(*
SPDX-FileCopyrightText: © 2026 Oleksandr Tiutyk <trofimich@gmail.com>
SPDX-License-Identifier: MIT
License: https://opensource.org/license/mit
*)

(*!
<summary>Orders WSTRING(255) values described by generic descriptors.</summary>
<description>
Non-null addresses must reference live WSTRING(255) storage. TypeClass and Size are not validated and no
numeric conversion is performed. Two null addresses compare equal; one null address sorts before a non-null
address. Uses native string comparison through the declared 255-character pointer type; descriptor Size does
not bound the read. Descriptors are passed by value; payload remains borrowed and is not modified, cloned,
released or retained. IsMemoryOwner does not affect comparison.
</description>
*)

FUNCTION_BLOCK WStringComparer EXTENDS TOF_Core.Object IMPLEMENTS TOF_Core.IComparer
VAR_STAT
	//! <summary>Class name shared by all instances of this function block.</summary>
	{attribute 'hide'} 
	_ClassName : STRING := __POUNAME();
END_VAR

{attribute 'monitoring' := 'call'}
PROPERTY ClassName : REFERENCE TO STRING
GET
ClassName REF= _ClassName;
END_GET
END_PROPERTY

(*!
<summary>Compares the first operand with the second using this ordering strategy.</summary>
<description>
Non-null addresses must reference live WSTRING(255) storage. TypeClass and Size are not validated and no
numeric conversion is performed. Two null addresses compare equal; one null address sorts before a non-null
address. Uses native string comparison through the declared 255-character pointer type; descriptor Size does
not bound the read. Descriptors are passed by value; payload remains borrowed and is not modified, cloned,
released or retained. IsMemoryOwner does not affect comparison. Descendants cannot replace this standard
ordering; implement IComparer separately for a different ordering strategy.
</description>
*)
//!<param name="first">First descriptor; referenced storage is borrowed for the call.</param>
//!<param name="second">Second descriptor; referenced storage is borrowed for the call.</param>
{attribute "object_name" := "Compare"}
METHOD FINAL Compare : TOF_Core.COMPARISON_RESULT
VAR_INPUT
	first : TOF_Core.GENERIC_VALUE;
	second : TOF_Core.GENERIC_VALUE;
END_VAR
VAR
	leftPointer : POINTER TO WSTRING(255); 
	rightPointer : POINTER TO WSTRING(255); 
END_VAR
IF first.Address = 0 AND_THEN second.Address = 0 THEN
	Compare := TOF_Core.COMPARISON_RESULT.FIRST_EQUAL_TO_SECOND;
	RETURN;
END_IF

IF first.Address = 0 THEN
	Compare := TOF_Core.COMPARISON_RESULT.FIRST_LESS_THAN_SECOND;
	RETURN;	
END_IF

IF second.Address = 0 THEN
	Compare := TOF_Core.COMPARISON_RESULT.FIRST_GREATER_THAN_SECOND;
	RETURN;	
END_IF

leftPointer := first.Address;
rightPointer := second.Address;

IF leftPointer^ < rightPointer^ THEN
	Compare := TOF_Core.COMPARISON_RESULT.FIRST_LESS_THAN_SECOND;
ELSIF leftPointer^ > rightPointer^ THEN
	Compare := TOF_Core.COMPARISON_RESULT.FIRST_GREATER_THAN_SECOND;
ELSE
	Compare := TOF_Core.COMPARISON_RESULT.FIRST_EQUAL_TO_SECOND;	
END_IF
END_METHOD

{attribute 'monitoring' := 'call'}
PROPERTY NamespaceName : REFERENCE TO STRING
GET
NamespaceName REF= CurrentNamespace.Name;
END_GET
END_PROPERTY

{attribute 'monitoring' := 'call'}
PROPERTY SelfSize : ULINT
GET
SelfSize := XSIZEOF(THIS^);
END_GET
END_PROPERTY

END_FUNCTION_BLOCK

(* stored: Version 1.1.0.1
   POU WStringComparer: Id {62ecc2ff-18fc-452f-b625-1d0f3cbba79c}, SpecialFunc None
   Property ClassName: Id {a81f1eb3-0ca7-4b4d-ae6f-d881ee745c52}
   Get Get: Id {d638f06b-8d02-44e3-bfd8-4933f9ab9a42}
   Method Compare: Id {e601d39a-f416-4f92-90c3-c07a65ebcb17}
   Property NamespaceName: Id {40543462-4099-4842-9c4b-f065b68e633d}
   Get Get: Id {9e6e185f-3d66-456d-a5c2-b0984348c06c}
   Property SelfSize: Id {d71f929e-eaa0-435c-83d2-409d58a515b6}
   Get Get: Id {0eaf5f05-5f99-40e9-80b5-39b36145a18f} *)
